FUNCTION_BLOCK SKILL_Join3 (* Ends a block of steps that run side by side: done when every branch is done; if one fails, the others are halted and the block fails. Technical: Ends a parallel block of 3 branches: DONE when all are done; on the first failure HALT to the others, then FAILED with its error once all have ended *)
  (* Standard: 61499-2 *)
  (* Version 0.1, 2026-09-28, Project contributors, AAU Smart Production Lab *)
  PACKAGE modlib;
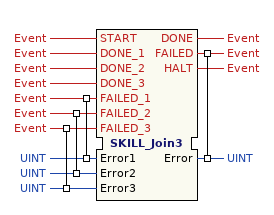
  EVENT_INPUT
    START; (* The parallel block starts: forget the last run *)
    DONE_1; (* Branch 1 is done *)
    DONE_2; (* Branch 2 is done *)
    DONE_3; (* Branch 3 is done *)
    FAILED_1 WITH Error1; (* Branch 1 failed (Error1) *)
    FAILED_2 WITH Error2; (* Branch 2 failed (Error2) *)
    FAILED_3 WITH Error3; (* Branch 3 failed (Error3) *)
  END_EVENT
  EVENT_OUTPUT
    DONE; (* Every branch is done *)
    FAILED WITH Error; (* A branch failed and every branch has ended (Error) *)
    HALT; (* A branch failed: stop the others *)
  END_EVENT
  VAR_INPUT
    Error1 : UINT; (* Error code of branch 1 *)
    Error2 : UINT; (* Error code of branch 2 *)
    Error3 : UINT; (* Error code of branch 3 *)
  END_VAR
  VAR_OUTPUT
    Error : UINT; (* Error code of the branch that failed first *)
  END_VAR
  VAR
    Ended1 : BOOL;
    Ended2 : BOOL;
    Ended3 : BOOL;
    AnyFailed : BOOL;
    First : UINT;
  END_VAR
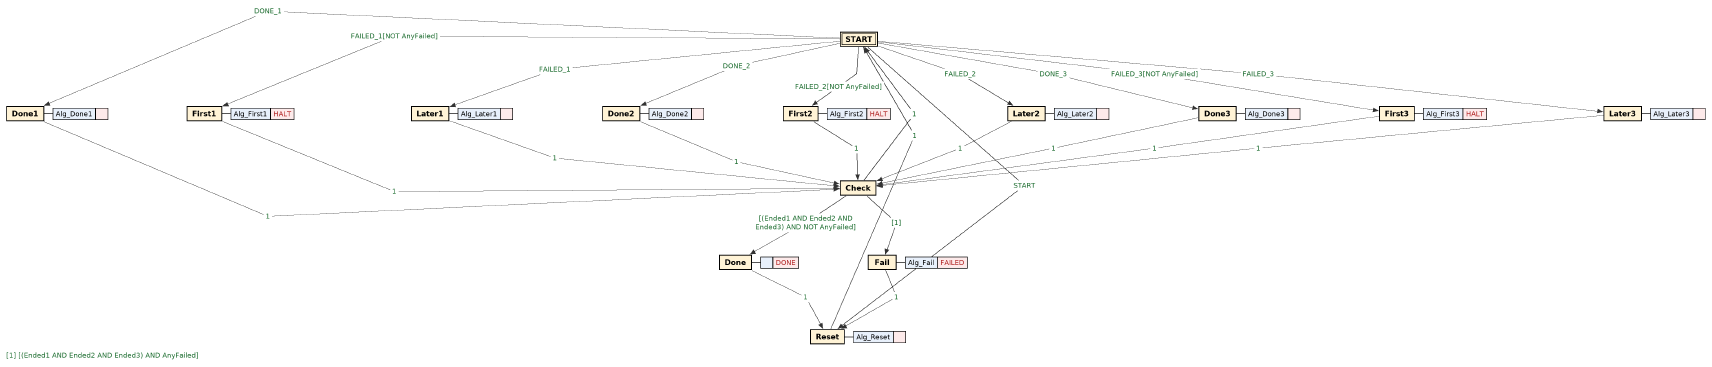
  EC_STATES
    START;
    Reset : Alg_Reset;
    Check;
    Done : -> DONE;
    Fail : Alg_Fail -> FAILED;
    Done1 : Alg_Done1;
    First1 : Alg_First1 -> HALT;
    Later1 : Alg_Later1;
    Done2 : Alg_Done2;
    First2 : Alg_First2 -> HALT;
    Later2 : Alg_Later2;
    Done3 : Alg_Done3;
    First3 : Alg_First3 -> HALT;
    Later3 : Alg_Later3;
  END_STATES
  EC_TRANSITIONS
    START TO Reset := START;
    Reset TO START := 1;
    START TO Done1 := DONE_1;
    START TO First1 := FAILED_1[NOT AnyFailed];
    START TO Later1 := FAILED_1;
    Done1 TO Check := 1;
    First1 TO Check := 1;
    Later1 TO Check := 1;
    START TO Done2 := DONE_2;
    START TO First2 := FAILED_2[NOT AnyFailed];
    START TO Later2 := FAILED_2;
    Done2 TO Check := 1;
    First2 TO Check := 1;
    Later2 TO Check := 1;
    START TO Done3 := DONE_3;
    START TO First3 := FAILED_3[NOT AnyFailed];
    START TO Later3 := FAILED_3;
    Done3 TO Check := 1;
    First3 TO Check := 1;
    Later3 TO Check := 1;
    Check TO Done := [(Ended1 AND Ended2 AND Ended3) AND NOT AnyFailed];
    Check TO Fail := [(Ended1 AND Ended2 AND Ended3) AND AnyFailed];
    Check TO START := 1;
    Done TO Reset := 1;
    Fail TO Reset := 1;
  END_TRANSITIONS
  ALGORITHM Alg_Reset IN ST:
Ended1 := FALSE; Ended2 := FALSE; Ended3 := FALSE; AnyFailed := FALSE;
  END_ALGORITHM
  ALGORITHM Alg_Fail IN ST:
Error := First;
  END_ALGORITHM
  ALGORITHM Alg_Done1 IN ST:
Ended1 := TRUE;
  END_ALGORITHM
  ALGORITHM Alg_First1 IN ST:
Ended1 := TRUE; AnyFailed := TRUE; First := Error1;
  END_ALGORITHM
  ALGORITHM Alg_Later1 IN ST:
Ended1 := TRUE;
  END_ALGORITHM
  ALGORITHM Alg_Done2 IN ST:
Ended2 := TRUE;
  END_ALGORITHM
  ALGORITHM Alg_First2 IN ST:
Ended2 := TRUE; AnyFailed := TRUE; First := Error2;
  END_ALGORITHM
  ALGORITHM Alg_Later2 IN ST:
Ended2 := TRUE;
  END_ALGORITHM
  ALGORITHM Alg_Done3 IN ST:
Ended3 := TRUE;
  END_ALGORITHM
  ALGORITHM Alg_First3 IN ST:
Ended3 := TRUE; AnyFailed := TRUE; First := Error3;
  END_ALGORITHM
  ALGORITHM Alg_Later3 IN ST:
Ended3 := TRUE;
  END_ALGORITHM
END_FUNCTION_BLOCK
